Staubli VAL3: moveTohome.pgx

program moveTohome()
begin
  call simulate:simulateHome()
end
